(* IEC 61131-3 sources: JingjiangArm/moonboxpro_arm_8.4/Application/Application/任务列表/Main_Task/套色调整, 11 files *)

(* ---- StAxisRapidAdjProf_H.st ---- *)
(*@CES
Name=StAxisRapidAdjProf_H
Type=Gvl
TypeGuid=2db5746d-d284-4425-9f7f-2663a34b0ebc
Guid=5051c563-c1c0-4e5b-a440-3f9f823cc70c
HasDeclaration=True
HasImplementation=False
*)
{DECLARATION}
TYPE StAxisRapidAdjProf_H :
STRUCT
	iIdxWr: INT; (* 索引-写 *)
	iIdxRd: INT; (* 索引-读 *)
	aiAdjustment: ARRAY [1..MAX_UNIT_NUM] OF INT; (* 快速调整量 *)
END_STRUCT
END_TYPE

{IMPLEMENTATION}

(* ---- StAxisRapidAdjProf_V.st ---- *)
(*@CES
Name=StAxisRapidAdjProf_V
Type=Gvl
TypeGuid=2db5746d-d284-4425-9f7f-2663a34b0ebc
Guid=880600c0-33b6-45cc-b2cb-0ddee2d5a314
HasDeclaration=True
HasImplementation=False
*)
{DECLARATION}
TYPE StAxisRapidAdjProf_V :
STRUCT
	iIdxWr: INT; (* 索引-写 *)
	iIdxRd: INT; (* 索引-读 *)
	adiAdjustment: ARRAY [1..MAX_UNIT_NUM] OF DINT; (* 快速调整量 *)
END_STRUCT
END_TYPE

{IMPLEMENTATION}

(* ---- KS_ClearRapidAdjValue_H.st ---- *)
(*@CES
Name=KS_ClearRapidAdjValue_H
Type=FunctionBlock
TypeGuid=6f9dac99-8de1-4efc-8465-68ac443b7d08
Guid=03f16b2d-6a59-44a0-871c-7df53a0c4716
HasDeclaration=True
HasImplementation=True
*)
{DECLARATION}
FUNCTION KS_ClearRapidAdjValue_H : INT(* 0:无错误/-1220:参数错误 *)
VAR_INPUT
	i_pastStAxisRapidAdjProf_H: POINTER TO ARRAY [1..MAX_UNIT_NUM] OF StAxisRapidAdjProf_H; (* 纵向快速对版 *)
	i_iUnitId: INT; (* 轴id *)
END_VAR
VAR
	iN: INT;
END_VAR

{IMPLEMENTATION}
IF i_pastStAxisRapidAdjProf_H<>0 AND
	i_iUnitId>=1 AND i_iUnitId<=MAX_UNIT_NUM THEN
	i_pastStAxisRapidAdjProf_H^[i_iUnitId].iIdxRd:= 1;
	i_pastStAxisRapidAdjProf_H^[i_iUnitId].iIdxWr:= 1;
	FOR iN:= 1 TO MAX_UNIT_NUM BY 1 DO
		i_pastStAxisRapidAdjProf_H^[i_iUnitId].aiAdjustment[iN]:= 0;
	END_FOR

ELSE
	KS_ClearRapidAdjValue_H:= -1220;
END_IF

KS_ClearRapidAdjValue_H:= 0;

(* ---- KS_ClearRapidAdjValue_V.st ---- *)
(*@CES
Name=KS_ClearRapidAdjValue_V
Type=FunctionBlock
TypeGuid=6f9dac99-8de1-4efc-8465-68ac443b7d08
Guid=1935351e-c560-4435-95d2-225c7524606b
HasDeclaration=True
HasImplementation=True
*)
{DECLARATION}
FUNCTION KS_ClearRapidAdjValue_V : INT(* 0:无错误/-1220:参数错误 *)
VAR_INPUT
	i_pastStAxisRapidAdjProf_V: POINTER TO ARRAY [1..MAX_UNIT_NUM] OF StAxisRapidAdjProf_V; (* 纵向快速对版 *)
	i_iUnitId: INT; (* 轴id *)
END_VAR
VAR
	iN: INT;
END_VAR

{IMPLEMENTATION}
IF i_pastStAxisRapidAdjProf_V<>0 AND
	i_iUnitId>=1 AND i_iUnitId<=MAX_UNIT_NUM THEN
	i_pastStAxisRapidAdjProf_V^[i_iUnitId].iIdxRd:= 1;
	i_pastStAxisRapidAdjProf_V^[i_iUnitId].iIdxWr:= 1;
	FOR iN:= 1 TO MAX_UNIT_NUM BY 1 DO
		i_pastStAxisRapidAdjProf_V^[i_iUnitId].adiAdjustment[iN]:= 0;
	END_FOR

ELSE
	KS_ClearRapidAdjValue_V:= -1220;
END_IF

KS_ClearRapidAdjValue_V:= 0;

(* ---- KS_ClearRegAdjValue.st ---- *)
(*@CES
Name=KS_ClearRegAdjValue
Type=FunctionBlock
TypeGuid=6f9dac99-8de1-4efc-8465-68ac443b7d08
Guid=35f4f50d-9372-488d-a3f0-1c615a8e6e33
HasDeclaration=True
HasImplementation=True
*)
{DECLARATION}
FUNCTION KS_ClearRegAdjValue : INT(* 0:无错误/-1220:参数错误 *)
VAR_INPUT
	i_pastStRegAdjMana: POINTER TO ARRAY [1..MAX_UNIT_NUM] OF StRegAdjMana; (* 单元调整量 *)
	i_iUnitId: INT; (* 轴id *)
END_VAR
VAR
	iN: INT;
END_VAR
{IMPLEMENTATION}
IF i_pastStRegAdjMana<>0 AND (*调整量结构体有效*)
	(i_iUnitId>=1 AND i_iUnitId<=MAX_UNIT_NUM) THEN (*轴id有效*)
	i_pastStRegAdjMana^[i_iUnitId].iIdxWr:= 1;
	i_pastStRegAdjMana^[i_iUnitId].iIdxRd:= 1;
	FOR iN:=1 TO GC_PU_MAX_NUM BY 1 DO
		i_pastStRegAdjMana^[i_iUnitId].aiAdj_V[iN]:= 0;
		i_pastStRegAdjMana^[i_iUnitId].aiAdj_H[iN]:= 0;
	END_FOR
	KS_ClearRegAdjValue:= 0;
ELSE
	KS_ClearRegAdjValue:= -1220;
END_IF

(* ---- KS_FetchRapidAdjValue_H.st ---- *)
(*@CES
Name=KS_FetchRapidAdjValue_H
Type=FunctionBlock
TypeGuid=6f9dac99-8de1-4efc-8465-68ac443b7d08
Guid=78ca29e0-c0c8-4d49-891a-0d1322be4c96
HasDeclaration=True
HasImplementation=True
*)
{DECLARATION}
FUNCTION KS_FetchRapidAdjValue_H : int
VAR_INPUT
	i_pastStAxisRapidAdjProf_H: POINTER TO ARRAY [1..MAX_UNIT_NUM] OF StAxisRapidAdjProf_H; (* 纵向快速对版| *)
	i_iUnitId: INT; (* 轴id| *)
	i_piValue: POINTER TO INT; (* 该轴对应的快速调版量| *)
END_VAR
VAR
	iResult: INT;
	iTempIndex: INT;
	iItemTotalNum: INT;
	iTemp: INT;
END_VAR

{IMPLEMENTATION}
iResult:= 0;
IF i_pastStAxisRapidAdjProf_H<>0 AND
	i_iUnitId>=1 AND i_iUnitId<=MAX_UNIT_NUM AND
	i_piValue<>0 THEN

	(*最大索引容量|*)
	iItemTotalNum:= SIZEOF(i_pastStAxisRapidAdjProf_H^[i_iUnitId].aiAdjustment)/SIZEOF(i_pastStAxisRapidAdjProf_H^[i_iUnitId].aiAdjustment[1]);

	IF i_pastStAxisRapidAdjProf_H^[i_iUnitId].iIdxRd<1 OR
		i_pastStAxisRapidAdjProf_H^[i_iUnitId].iIdxRd>iItemTotalNum OR
		i_pastStAxisRapidAdjProf_H^[i_iUnitId].iIdxWr<1 OR
		i_pastStAxisRapidAdjProf_H^[i_iUnitId].iIdxWr>iItemTotalNum THEN
		(*如果索引异常就全部清空不处理|*)
		i_pastStAxisRapidAdjProf_H^[i_iUnitId].iIdxRd:= 1;
		i_pastStAxisRapidAdjProf_H^[i_iUnitId].iIdxWr:= 1;
		iResult:= 1220;
	ELSIF i_pastStAxisRapidAdjProf_H^[i_iUnitId].iIdxRd<>i_pastStAxisRapidAdjProf_H^[i_iUnitId].iIdxWr THEN
		(*有数据需要读取|*)
		(*写入出口位置|*)
		i_piValue^:= i_pastStAxisRapidAdjProf_H^[i_iUnitId].aiAdjustment[i_pastStAxisRapidAdjProf_H^[i_iUnitId].iIdxRd];

		(*下次读取的位置|*)
		iTempIndex:= i_pastStAxisRapidAdjProf_H^[i_iUnitId].iIdxRd+1;
		IF iTempIndex>iItemTotalNum THEN
			iTempIndex:= iTempIndex-iItemTotalNum;
		END_IF
		i_pastStAxisRapidAdjProf_H^[i_iUnitId].iIdxRd:= iTempIndex;
	ELSE
		(*没有新数据|*)
		iResult:= 1221;
	END_IF
ELSE
	iResult:= -1220;
END_IF

KS_FetchRapidAdjValue_H:= iResult;

(* ---- KS_FetchRapidAdjValue_V.st ---- *)
(*@CES
Name=KS_FetchRapidAdjValue_V
Type=FunctionBlock
TypeGuid=6f9dac99-8de1-4efc-8465-68ac443b7d08
Guid=43d9692c-d0f7-4421-a5e4-fec02edd6bb4
HasDeclaration=True
HasImplementation=True
*)
{DECLARATION}
FUNCTION KS_FetchRapidAdjValue_V : INT (* -1220:参数无效; 1220:读写索引无效(从头置位);1221:没有新的值; 0:无错误 *)
VAR_INPUT
	i_pastStAxisRapidAdjProf_V: POINTER TO ARRAY [1..MAX_UNIT_NUM] OF StAxisRapidAdjProf_V; (* 纵向快速对版 *)
	i_iUnitId: INT; (* 轴id *)
	i_pdiValue: POINTER TO DINT; (* 该轴对应的快速调版量 *)
END_VAR
VAR
	iResult: INT;
	iTempIndex: INT;
	iItemTotalNum: INT;
	diTemp: DINT;
END_VAR

{IMPLEMENTATION}
iResult:= 0;
IF i_pastStAxisRapidAdjProf_V<>0 AND
	i_iUnitId>=1 AND i_iUnitId<=MAX_UNIT_NUM AND
	i_pdiValue<>0 THEN

	(* 最大索引容量 *)
	iItemTotalNum:= SIZEOF(i_pastStAxisRapidAdjProf_V^[i_iUnitId].adiAdjustment)/SIZEOF(i_pastStAxisRapidAdjProf_V^[i_iUnitId].adiAdjustment[1]);

	IF i_pastStAxisRapidAdjProf_V^[i_iUnitId].iIdxRd<1 OR
		i_pastStAxisRapidAdjProf_V^[i_iUnitId].iIdxRd>iItemTotalNum OR
		i_pastStAxisRapidAdjProf_V^[i_iUnitId].iIdxWr<1 OR
		i_pastStAxisRapidAdjProf_V^[i_iUnitId].iIdxWr>iItemTotalNum THEN
		(* 如果索引异常就全部清空不处理 *)
		i_pastStAxisRapidAdjProf_V^[i_iUnitId].iIdxRd:= 1;
		i_pastStAxisRapidAdjProf_V^[i_iUnitId].iIdxWr:= 1;
		iResult:= 1220;
	ELSIF i_pastStAxisRapidAdjProf_V^[i_iUnitId].iIdxRd<>i_pastStAxisRapidAdjProf_V^[i_iUnitId].iIdxWr THEN
		(* 有数据需要读取 *)
		(* 写入出口位置 *)
		i_pdiValue^:= i_pastStAxisRapidAdjProf_V^[i_iUnitId].adiAdjustment[i_pastStAxisRapidAdjProf_V^[i_iUnitId].iIdxRd];

		(* 下次读取的位置 *)
		iTempIndex:= i_pastStAxisRapidAdjProf_V^[i_iUnitId].iIdxRd+1;
		IF iTempIndex>iItemTotalNum THEN
			iTempIndex:= iTempIndex-iItemTotalNum;
		END_IF
		i_pastStAxisRapidAdjProf_V^[i_iUnitId].iIdxRd:= iTempIndex;
	ELSE
		(* 没有新数据 *)
		iResult:= 1221;
	END_IF
ELSE
	iResult:= -1220;
END_IF

KS_FetchRapidAdjValue_V:= iResult;

(* ---- KS_FetchRegAdjValue.st ---- *)
(*@CES
Name=KS_FetchRegAdjValue
Type=FunctionBlock
TypeGuid=6f9dac99-8de1-4efc-8465-68ac443b7d08
Guid=1dd2d585-55d6-4e53-9602-3ae775b26755
HasDeclaration=True
HasImplementation=True
*)
{DECLARATION}
FUNCTION KS_FetchRegAdjValue : INT (* -1220:参数无效/1220:操作指针无效(并作复位处理)/0:无错误 *)
VAR_INPUT
	i_pastStRegAdjMana: POINTER TO ARRAY [1..MAX_UNIT_NUM] OF StRegAdjMana; (* 单元调整量 *)
	i_iUnitId: INT; (* 轴id *)
	i_piAdj_V: POINTER TO INT; (* 用以返回纵向调整量 *)
	i_piAdj_H: POINTER TO INT; (* 用以返回横向调整量 *)
END_VAR
VAR
	iResult: INT;
	iItemTotalNum: INT; (* 数据总量 *)
	iTmpValue: INT;
END_VAR
{IMPLEMENTATION}
iResult:= 0;
IF i_pastStRegAdjMana<>0 AND (*调整量结构体有效*)
	(i_iUnitId>=1 AND i_iUnitId<=MAX_UNIT_NUM) AND (*轴id有效*)
	(i_piAdj_V<>0 AND i_piAdj_H<>0) THEN (*返回地址有效*)
	iItemTotalNum:= SIZEOF(i_pastStRegAdjMana^[i_iUnitId].aiAdj_V)/SIZEOF(i_pastStRegAdjMana^[i_iUnitId].aiAdj_V[1]);
	IF (i_pastStRegAdjMana^[i_iUnitId].iIdxWr<1 OR i_pastStRegAdjMana^[i_iUnitId].iIdxWr>iItemTotalNum) OR
		(i_pastStRegAdjMana^[i_iUnitId].iIdxRd<1 OR i_pastStRegAdjMana^[i_iUnitId].iIdxRd>iItemTotalNum) THEN
		(*索引无效*)
		i_pastStRegAdjMana^[i_iUnitId].iIdxRd:= 1;
		i_pastStRegAdjMana^[i_iUnitId].iIdxWr:= 1;
		iResult:= 1220;
	ELSIF i_pastStRegAdjMana^[i_iUnitId].iIdxWr<>i_pastStRegAdjMana^[i_iUnitId].iIdxRd THEN
		(*队列不齐*)
		i_piAdj_V^:= i_pastStRegAdjMana^[i_iUnitId].aiAdj_V[i_pastStRegAdjMana^[i_iUnitId].iIdxRd];
		i_piAdj_H^:= i_pastStRegAdjMana^[i_iUnitId].aiAdj_H[i_pastStRegAdjMana^[i_iUnitId].iIdxRd];

		(*定位下次要访问的位置*)
		iTmpValue:= i_pastStRegAdjMana^[i_iUnitId].iIdxRd+1;
		IF iTmpValue>iItemTotalNum THEN
			iTmpValue:= iTmpValue-iItemTotalNum;
		END_IF
		i_pastStRegAdjMana^[i_iUnitId].iIdxRd:= iTmpValue;
	ELSE(*2018.8.21.202154\修复bug\基本可以怀疑是这里的问题了\折腾了好多天|*)
		(*忘记else分支最后造成返回值为默认的0|这样之前的值会被重复使用|造成调整量量增|*)
		iResult:= 1221;
	END_IF
ELSE
	iResult:= -1220;
END_IF

KS_FetchRegAdjValue:= iResult;

(* ---- KS_PushRapidAdjValue_H.st ---- *)
(*@CES
Name=KS_PushRapidAdjValue_H
Type=FunctionBlock
TypeGuid=6f9dac99-8de1-4efc-8465-68ac443b7d08
Guid=f4c3ad13-cefe-4439-a936-6639860b4e75
HasDeclaration=True
HasImplementation=True
*)
{DECLARATION}
FUNCTION KS_PushRapidAdjValue_H : INT(*0:无错误; -1220:参数错误|*)
VAR_INPUT
	i_pastStAxisRapidAdjProf_H: POINTER TO ARRAY [1..MAX_UNIT_NUM] OF StAxisRapidAdjProf_H; (* 纵向快速对版| *)
	i_iUnitId: INT; (* 轴id| *)
	i_iValue: INT; (* 提交的数据 *)
END_VAR
VAR
	iResult: INT;
	iTempIndex: INT;
	iItemTotalNum: INT;
END_VAR

{IMPLEMENTATION}
iResult:= 0;
IF i_pastStAxisRapidAdjProf_H<>0 AND
	i_iUnitId>=1 AND i_iUnitId<=MAX_UNIT_NUM AND
	i_iValue<>0 THEN

	(*先算出最大容量|*)
	iItemTotalNum:= SIZEOF(i_pastStAxisRapidAdjProf_H^[i_iUnitId].aiAdjustment)/SIZEOF(i_pastStAxisRapidAdjProf_H^[i_iUnitId].aiAdjustment[1]);

	(*如果索引超限|默认清空从头开始|*)
	IF i_pastStAxisRapidAdjProf_H^[i_iUnitId].iIdxRd<1 OR(*读索引超限|*)
		i_pastStAxisRapidAdjProf_H^[i_iUnitId].iIdxRd>iItemTotalNum OR
		i_pastStAxisRapidAdjProf_H^[i_iUnitId].iIdxWr<1 OR(*写索引超限|*)
		i_pastStAxisRapidAdjProf_H^[i_iUnitId].iIdxWr>iItemTotalNum THEN
		i_pastStAxisRapidAdjProf_H^[i_iUnitId].iIdxRd:= 1;
		i_pastStAxisRapidAdjProf_H^[i_iUnitId].iIdxWr:= 1;
	END_IF

	(*写入新值|*)
	i_pastStAxisRapidAdjProf_H^[i_iUnitId].aiAdjustment[i_pastStAxisRapidAdjProf_H^[i_iUnitId].iIdxWr]:= i_iValue;

	(*定位到下次写入位置|*)
	iTempIndex:= i_pastStAxisRapidAdjProf_H^[i_iUnitId].iIdxWr+1;
	IF iTempIndex>iItemTotalNum THEN
		iTempIndex:= iTempIndex-iItemTotalNum;
	END_IF
	i_pastStAxisRapidAdjProf_H^[i_iUnitId].iIdxWr:= iTempIndex;
ELSE
	iResult:= -1220;
END_IF

KS_PushRapidAdjValue_H:= iResult;

(* ---- KS_PushRapidAdjValue_V.st ---- *)
(*@CES
Name=KS_PushRapidAdjValue_V
Type=FunctionBlock
TypeGuid=6f9dac99-8de1-4efc-8465-68ac443b7d08
Guid=78c765c0-3731-4952-bfd4-57dc02a59b2a
HasDeclaration=True
HasImplementation=True
*)
{DECLARATION}
FUNCTION KS_PushRapidAdjValue_V : INT(*0:无错误; -1220:参数错误|*)
VAR
	iResult: INT;
	iTempIndex: INT;
	iItemTotalNum: INT;
END_VAR
VAR_INPUT
	i_pastStAxisRapidAdjProf_V: POINTER TO ARRAY [1..MAX_UNIT_NUM] OF StAxisRapidAdjProf_V; (* 纵向快速对版| *)
	i_iUnitId: INT; (* 轴id| *)
	i_diValue: DINT; (* 提交的数据 *)
END_VAR

{IMPLEMENTATION}
iResult:= 0;
IF i_pastStAxisRapidAdjProf_V<>0 AND
	i_iUnitId>=1 AND i_iUnitId<=MAX_UNIT_NUM AND
	i_diValue<>0 THEN

	(*先算出最大容量|*)
	iItemTotalNum:= SIZEOF(i_pastStAxisRapidAdjProf_V^[i_iUnitId].adiAdjustment)/SIZEOF(i_pastStAxisRapidAdjProf_V^[i_iUnitId].adiAdjustment[1]);

	(*如果索引超限|默认清空从头开始|*)
	IF i_pastStAxisRapidAdjProf_V^[i_iUnitId].iIdxRd<1 OR(*读索引超限|*)
		i_pastStAxisRapidAdjProf_V^[i_iUnitId].iIdxRd>iItemTotalNum OR
		i_pastStAxisRapidAdjProf_V^[i_iUnitId].iIdxWr<1 OR(*写索引超限|*)
		i_pastStAxisRapidAdjProf_V^[i_iUnitId].iIdxWr>iItemTotalNum THEN
		i_pastStAxisRapidAdjProf_V^[i_iUnitId].iIdxRd:= 1;
		i_pastStAxisRapidAdjProf_V^[i_iUnitId].iIdxWr:= 1;
	END_IF

	(*写入新值|*)
	i_pastStAxisRapidAdjProf_V^[i_iUnitId].adiAdjustment[i_pastStAxisRapidAdjProf_V^[i_iUnitId].iIdxWr]:= i_diValue;

	(*定位到下次写入位置|*)
	iTempIndex:= i_pastStAxisRapidAdjProf_V^[i_iUnitId].iIdxWr+1;
	IF iTempIndex>iItemTotalNum THEN
		iTempIndex:= iTempIndex-iItemTotalNum;
	END_IF
	i_pastStAxisRapidAdjProf_V^[i_iUnitId].iIdxWr:= iTempIndex;
ELSE
	iResult:= -1220;
END_IF

KS_PushRapidAdjValue_V:= iResult;

(* ---- KS_PushRegAdjValue.st ---- *)
(*@CES
Name=KS_PushRegAdjValue
Type=FunctionBlock
TypeGuid=6f9dac99-8de1-4efc-8465-68ac443b7d08
Guid=5b088804-504f-459b-bb64-be78c2ffc3f4
HasDeclaration=True
HasImplementation=True
*)
{DECLARATION}
FUNCTION KS_PushRegAdjValue : INT(* 0:无错误/-1220:参数错误 *)
VAR_INPUT
	i_pastStRegAdjMana: POINTER TO ARRAY [1..MAX_UNIT_NUM] OF StRegAdjMana; (* 单元调整量 *)
	i_iUnitId: INT; (* 轴id *)
	i_iAdj_V: INT; (* 纵向调整量 *)
	i_iAdj_H: INT; (* 横向调整量 *)
END_VAR
VAR
	iItemTotalNum: INT; (* 数据总量 *)
	iTmpValue: INT;
END_VAR
{IMPLEMENTATION}
IF i_pastStRegAdjMana<>0 AND (*调整量结构体有效*)
	(i_iUnitId>=1 AND i_iUnitId<=MAX_UNIT_NUM) THEN (*轴id有效*)
	iItemTotalNum:= SIZEOF(i_pastStRegAdjMana^[i_iUnitId].aiAdj_V)/SIZEOF(i_pastStRegAdjMana^[i_iUnitId].aiAdj_V[1]);
	IF (i_pastStRegAdjMana^[i_iUnitId].iIdxWr<1 OR i_pastStRegAdjMana^[i_iUnitId].iIdxWr>iItemTotalNum) OR
		(i_pastStRegAdjMana^[i_iUnitId].iIdxRd<1 OR i_pastStRegAdjMana^[i_iUnitId].iIdxRd>iItemTotalNum) THEN
		i_pastStRegAdjMana^[i_iUnitId].iIdxRd:= 1;
		i_pastStRegAdjMana^[i_iUnitId].iIdxWr:= 1;
	END_IF

	i_pastStRegAdjMana^[i_iUnitId].aiAdj_V[i_pastStRegAdjMana^[i_iUnitId].iIdxWr]:= i_iAdj_V; (*写入纵向调整量*)
	i_pastStRegAdjMana^[i_iUnitId].aiAdj_H[i_pastStRegAdjMana^[i_iUnitId].iIdxWr]:= i_iAdj_H; (*写入横向调整量*)

	(*处理下一次要写入数据的位置
	.由于Push和Fetch最终会在两个优先级不同的任务中执行
	.每个函数调用时都会先检查索引是否有效
	.所以为了保证变量的原子态操作
	.所以把+1和判断放在临时变量中操作
	*)
	iTmpValue:= i_pastStRegAdjMana^[i_iUnitId].iIdxWr+1;
	IF iTmpValue>iItemTotalNum THEN
		iTmpValue:= iTmpValue-iItemTotalNum;
	END_IF
	i_pastStRegAdjMana^[i_iUnitId].iIdxWr:= iTmpValue;

	KS_PushRegAdjValue:= 0;
ELSE
	KS_PushRegAdjValue:= -1220;
END_IF
